{attribute 'no_assign'}
FUNCTION_BLOCK FB_DO_WTURBINE_LD0_WTUR1_DmdWSpt_val EXTENDS FB_AcsiCommonControllableDataClass
VAR_INPUT
	origin: FB_AcsiDATypeOriginator := (Fc:=ACSI_FC_MX, bLinkResult:=THIS^.AddDataToContainer(ipData:=origin));
	mxVal: FB_AcsiDATypeAnalogueValue := (Fc:=ACSI_FC_MX, TrgOp:=ACSI_TrgOp_dchg, i:=(bPresence:=FALSE), bLinkResult:=THIS^.AddDataToContainer(ipData:=mxVal));
	q: FB_AcsiDATypeQuality := (Fc:=ACSI_FC_MX, TrgOp:=ACSI_TrgOp_qchg, bLinkResult:=THIS^.AddDataToContainer(ipData:=q));
	t: FB_AcsiDATypeTimeStamp := (Fc:=ACSI_FC_MX, bLinkResult:=THIS^.AddDataToContainer(ipData:=t));
	ctlModel: FB_AcsiDATypeCtlModels := (Fc:=ACSI_FC_CF, TrgOp:=ACSI_TrgOp_dchg, eValue:=E_AcsiCtlModels.DirectWithNormalSecurity, bLinkResult:=THIS^.AddDataToContainer(ipData:=ctlModel));
	Oper: FB_AcsiCDC_Oper_AnalogueValue := (Fc:=ACSI_FC_CO, ctlVal:=(i:=(bPresence:=FALSE)), bLinkResult:=THIS^.AddDataToContainer(ipData:=Oper));
	SBO: FB_AcsiCDC_SBO := (Fc:=ACSI_FC_CO, bLinkResult:=THIS^.AddDataToContainer(ipData:=SBO));
	Cancel: FB_AcsiCDC_Cancel_AnalogueValue := (Fc:=ACSI_FC_CO, ctlVal:=(i:=(bPresence:=FALSE)), bLinkResult:=THIS^.AddDataToContainer(ipData:=Cancel));
	
	fbControl: FB_DirectControl := (ipCtrl:=THIS^.AddServerJob(ipEvent:=fbControl, ipCompletion:=fbControl));
// 	fbControl: FB_SboControl := (ipCtrl:=THIS^.AddServerJob(ipEvent:=fbControl, ipCompletion:=fbControl));
END_VAR
VAR
END_VAR

END_FUNCTION_BLOCK

(* stored: Version 1.1.0.1
   POU FB_DO_WTURBINE_LD0_WTUR1_DmdWSpt_val: Id {f1c47eca-556f-4a9e-8ad0-6c3dec6ae599}, SpecialFunc None *)
